TYPE "DT_ALM_ALL"
VERSION : 0.1
   STRUCT
      TURBINE : "DT_ALM_SYSTEM_TURBINE";
      HPU_PUMPS : "DT_ALM_SYSTEM_HPU_PUMPS";
      HPU : "DT_ALM_SYSTEM_HPU";
      WATERWAY : "DT_ALM_SYSTEM_WATERWAY";
      GEN_TEMP_WIND : "DT_ALM_SYSTEM_GEN_TEMP_WIND";
      GEN_BEAR_AND_AIR : "DT_ALM_SYSTEM_GEN_BEAR_AND_AIR";
      GEN_SPEED_WH_AND_VIB : "DT_ALM_SYSTEM_GEN_SPEED_WH_AND_VIB";
      GEN_OTHER_ALM : "DT_ALM_SYSTEM_GEN_OTHER_ALM";
      UNIT_TRAFO : "DT_ALM_SYSTEM_UNIT_TRAFO";
      AUX_TRAFO_AND_DIESEL : "DT_ALM_SYSTEM_AUX_TRAFO_AND_DIESEL";
      EXC_AND_SYNC : "DT_ALM_SYSTEM_EXC_AND_SYNC";
      PROT_AND_AUTO_MODE : "DT_ALM_SYSTEM_PROT_AND_AUTO_MODE";
      CTRL_AND_COMM_1 : "DT_ALM_SYSTEM_CTRL_AND_COMM_1";
      CTRL_AND_COMM_2 : "DT_ALM_SYSTEM_CTRL_AND_COMM_2";
      GEN_CUB_AND_OTHER : "DT_ALM_SYSTEM_GEN_CUB_AND_OTHER";
      AUX_AC_DC_1 : "DT_ALM_SYSTEM_AUX_AC_DC_1";
      AUX_AC_DC_2 : "DT_ALM_SYSTEM_AUX_AC_DC_2";
      SN_LINE : "DT_ALM_SYSTEM_SN_LINE";
      SN_GEN_AND_MEAS : "DT_ALM_SYSTEM_SN_GEN_AND_MEAS";
      SN_AUX_TRAFO_AND_GND : "DT_ALM_SYSTEM_SN_AUX_TRAFO_AND_GND";
      INTAKE : "DT_ALM_SYSTEM_INTAKE";
      CWS : "DT_ALM_SYSTEM_CWS";
      LOU : "DT_ALM_SYSTEM_LOU";
      DWS_AND_DRAIN : "DT_ALM_SYSTEM_DWS_AND_DRAIN";
      GEN_PROT_ALM : "DT_ALM_SYSTEM_SPARE_24";
      TRAFO_PROT_ALM : "DT_ALM_SYSTEM_SPARE_25";
      SPARE_26 : "DT_ALM_SYSTEM_SPARE_26";
      SPARE_27 : "DT_ALM_SYSTEM_SPARE_27";
      SPARE_28 : "DT_ALM_SYSTEM_SPARE_28";
      SPARE_29 : "DT_ALM_SYSTEM_SPARE_29";
      SPARE_30 : "DT_ALM_SYSTEM_SPARE_30";
   END_STRUCT;

END_TYPE

